// TIA Portal V20 export
DATA_BLOCK "T10_Resultado"   // DB47901
{ S7_Optimized_Access := 'TRUE' }
AUTHOR : IA
FAMILY : PRUEBA
VERSION : 0.1
// Tanda 4B: comunicación en marcha
// stored: AutoNumber false
   VAR
      S_TSEND_C_TRCV_C : Bool;   // TSEND_C → TRCV_C (puerto 2001): llegan los 4 bytes
      S_TCON_TSEND_TRCV : Bool;   // TCON ×2 + TSEND → TRCV (puerto 2002): llegan los 4 bytes
      S_TDISCON : Bool;   // TDISCON cierra la conexión cliente
      S_Modbus : Bool;   // MB_CLIENT lee 2 registros de MB_SERVER (puerto 502)
      Vida : DInt;   // Sube cada ciclo
      OK : Int;   // Correctas
      Total : Int := 4;   // Pruebas
      Todo_OK : Bool;   // Todas correctas
   END_VAR
BEGIN
END_DATA_BLOCK
